Staubli VAL3: MainLongProg.pjx

--- MainLongProg.pjx ---
Parameters version=s7.3.1 stackSize=5000 millimeterUnit=true
Program file=loadNextOne.pgx
Program file=start.pgx
Program file=stop.pgx
Data file=MainLongProg.dtx
Library alias=prog path=./LongProg/LongProg.pjx
Library alias=prog_swap path=./LongProg/LongProg.pjx
Library alias=tooldata path=saveChangeTool

--- MainLongProg.dtx ---
mdesc mNomSpeed
frame fFrame1 = {x=1234.570, y=-98.765, z=50.500, rx=-0.000, ry=0.000, rz=30.000, fatherId=world[0]}
dio Input[16]
  [0] = {link=BasicIO-1\%I0}
  [1] = {link=BasicIO-1\%I1}
  [2] = {link=BasicIO-1\%I2}
  [3] = {link=BasicIO-1\%I3}
  [4] = {link=BasicIO-1\%I4}
  [5] = {link=BasicIO-1\%I5}
  [6] = {link=BasicIO-1\%I6}
  [7] = {link=BasicIO-1\%I7}
  [8] = {link=BasicIO-1\%I8}
  [9] = {link=BasicIO-1\%I9}
  [10] = {link=BasicIO-1\%I10}
  [11] = {link=BasicIO-1\%I11}
  [12] = {link=BasicIO-1\%I12}
  [13] = {link=BasicIO-1\%I13}
  [14] = {link=BasicIO-1\%I14}
  [15] = {link=BasicIO-1\%I15}
dio Output[16]
  [0] = {link=BasicIO-1\%Q0}
  [1] = {link=BasicIO-1\%Q1}
  [2] = {link=BasicIO-1\%Q2}
  [3] = {link=BasicIO-1\%Q3}
  [4] = {link=BasicIO-1\%Q4}
  [5] = {link=BasicIO-1\%Q5}
  [6] = {link=BasicIO-1\%Q6}
  [7] = {link=BasicIO-1\%Q7}
  [8] = {link=BasicIO-1\%Q8}
  [9] = {link=BasicIO-1\%Q9}
  [10] = {link=BasicIO-1\%Q10}
  [11] = {link=BasicIO-1\%Q11}
  [12] = {link=BasicIO-1\%Q12}
  [13] = {link=BasicIO-1\%Q13}
  [14] = {link=BasicIO-1\%Q14}
  [15] = {link=BasicIO-1\%Q15}
tool tCurrentTool = {x=10.000, y=20.000, z=150.000, rx=-0.000, ry=0.000, rz=-0.000, fatherId=flange[0], ioLink=ValveIO/valve1}
mdesc mCurrentSpeed
pointRs pPointRs = {fatherId=fFrame1[0]}
pointRs pPointRs2 = {fatherId=fFrame1[0]}

--- start.pgx ---
public program start()
begin
  if prog:libLoad("./LongProg")!=0
    logMsg("Error Loading RoboDK library")
    popUpMsg("Error Loading RoboDK library")
  endIf
  wait(taskStatus("loading")==-1)
  taskCreate "loading",10,loadNextOne("./LongProg2")
  call prog:start()

  if prog:libLoad("./LongProg2")!=0
    logMsg("Error Loading RoboDK library")
    popUpMsg("Error Loading RoboDK library")
  endIf
  wait(taskStatus("loading")==-1)
  taskCreate "loading",10,loadNextOne("./LongProg3")
  call prog:start()

  if prog:libLoad("./LongProg3")!=0
    logMsg("Error Loading RoboDK library")
    popUpMsg("Error Loading RoboDK library")
  endIf
  wait(taskStatus("loading")==-1)
  call prog:start()


end

--- loadNextOne.pgx ---
program loadNextOne(string x_sName)
begin
  prog_swap:libLoad(x_sName)
end

--- stop.pgx ---
program stop()
begin
end
